(* IEC 61131-3 sources: codesys-framework/txt/application/ToDo/Warnings and Alarms, 15 files *)

(* ---- E_EventLevels.dut.st ---- *)
{attribute 'qualified_only'}
{attribute 'strict'}
TYPE E_EventLevels :
(
	Invalid := 0,
	NotApplicable := 1,
	Success := 5,
	EventIsInformational := 10,
	EventIsWarning_NotUrgent := 20,
	EventIsWarning_Urgent := 21,
	EventIsAlarm_OnlyLogLevel := 40,
	EventIsAlarm_OperatorLevel := 41,
	EventIsAlarm_SupervisorLevel := 42
);
END_TYPE

(* ---- SC_EventConfig.dut.st ---- *)
TYPE SC_EventConfig :
STRUCT
	udiEventID 						: UDINT;
	eSubMachine 					: INT;
	xEventIsDisabled 				: BOOL := FALSE;
	eEventLevel_InCaseOfWarning 	: E_EventLevels;
	eEventLevel_InCaseOfAlarm 		: E_EventLevels;
END_STRUCT
END_TYPE

(* ---- SC_EventHandler.dut.st ---- *)
TYPE SC_EventHandler :
STRUCT
	scEventConfig 					: SC_EventConfig;
	eEventLevel 					: E_EventLevels;
	xEvent_WarningIsActive 			: BOOL;
	xEvent_AlarmIsActive 			: BOOL;
	xEvent_WarningInsertedInLog 	: BOOL;
	xEvent_AlarmInsertedInLog 		: BOOL;
END_STRUCT
END_TYPE

(* ---- F_Event_InsertInLog.pou.st ---- *)
FUNCTION F_Event_InsertInLog : BOOL
VAR_INPUT
	eSubMachine 			: INT;
	w 						: WORD;
	udiEventID 				: UDINT;
	eEventLevel 			: E_EventLevels;
	asEventPayload 			: ARRAY [1..cHYP_MAX_PAYLOADFIELDS] OF STRING;
END_VAR
VAR
	_scEventForHyperion 	: SC_Hyperion_EventStruct;
END_VAR

// --- BEGIN IMPLEMENTATION ---

IF eSubMachine = E_SubMachines.YarnStorage THEN
	audiYSEventCounter[w] := audiYSEventCounter[w] + 1;
	_scEventForHyperion.Counter := audiYSEventCounter[w];

	IF audiYSEventCounter[w] >= 4294967295 THEN
		audiYSEventCounter[w] := 0;
	END_IF

ELSIF eSubMachine = E_SubMachines.CardBoardStorage THEN
	udiCSEventCounter := udiCSEventCounter + 1;
	_scEventForHyperion.Counter := udiCSEventCounter;

	IF udiCSEventCounter >= 4294967295 THEN
		udiCSEventCounter := 0;
	END_IF

ELSE
	udiFREventCounter := udiFREventCounter + 1;
	_scEventForHyperion.Counter := udiFREventCounter;

	IF udiFREventCounter >= 4294967295 THEN
		udiFREventCounter := 0;
	END_IF

END_IF

_scEventForHyperion.Identification := udiEventID;

(*
IF eSubMachine = E_SubMachines.Creel THEN
	audiCLEventCounter[w] := audiCLEventCounter[w] + 1;
	_scEventForHyperion.Counter := audiCLEventCounter[w];
ELSIF eSubMachine = E_SubMachines.CreelRobot THEN
	audiCREventCounter[w] := audiCREventCounter[w] + 1;
	_scEventForHyperion.Counter := audiCREventCounter[w];
ELSIF eSubMachine = E_SubMachines.CreelConveyor THEN
	audiCCEventCounter[w] := audiCCEventCounter[w] + 1;
	_scEventForHyperion.Counter := audiCCEventCounter[w];
ELSIF eSubMachine = E_SubMachines.YarnConsumer THEN
	audiHSEventCounter[w] := audiHSEventCounter[w] + 1;
	_scEventForHyperion.Counter := audiHSEventCounter[w];
ELSE
	udiCUEventCounter := udiCUEventCounter + 1;
	_scEventForHyperion.Counter := udiCUEventCounter;
END_IF
*)

_scEventForHyperion.Identification := udiEventID;

// Create Hyperion Event Struct
CASE (eEventLevel) OF
	E_EventLevels.EventIsInformational : _scEventForHyperion.Level := cHYP_LEVEL_INFORMATIONAL;
	E_EventLevels.Success : _scEventForHyperion.Level := cHYP_LEVEL_BOOKMARK;
	E_EventLevels.EventIsWarning_NotUrgent : _scEventForHyperion.Level := cHYP_LEVEL_WARNING;
	E_EventLevels.EventIsWarning_Urgent : _scEventForHyperion.Level := cHYP_LEVEL_WARNING;
	E_EventLevels.EventIsAlarm_OnlyLogLevel : _scEventForHyperion.Level := cHYP_LEVEL_ERROR;
	E_EventLevels.EventIsAlarm_OperatorLevel : _scEventForHyperion.Level := cHYP_LEVEL_ERROR;
	E_EventLevels.EventIsAlarm_SupervisorLevel : _scEventForHyperion.Level := cHYP_LEVEL_ERROR;
END_CASE

// _scEventForHyperion.TimeStamp := sTimeStamp_Local_AsString;
_scEventForHyperion.TimeStamp := sTimeStamp_UTC_AsString;
_scEventForHyperion.PayLoad := F_HyperionCreatePayloadString (asEventPayload := asEventPayload);

// Insert in local eventbuffer
IF eSubMachine = E_SubMachines.YarnStorage THEN
	audiYSLocalEventPointer[w] := audiYSLocalEventPointer[w] + 1;
	IF audiYSLocalEventPointer[w] > cMaxLocalEvents THEN
		audiYSLocalEventPointer[w] := 1;
	END_IF
	aascYSLocalEventList[w][audiYSLocalEventPointer[w]].udiEventID := udiEventID;
	aascYSLocalEventList[w][audiYSLocalEventPointer[w]].eEventLevel := eEventLevel;

ELSE
	udiFRLocalEventPointer := udiFRLocalEventPointer + 1;
	IF udiFRLocalEventPointer > cMaxLocalEvents THEN
		udiFRLocalEventPointer := 1;
	END_IF
	ascFRLocalEventList[udiFRLocalEventPointer].udiEventID := udiEventID;
	ascFRLocalEventList[udiFRLocalEventPointer].eEventLevel := eEventLevel;
END_IF

// Insert in Hyperion eventbuffer
IF eSubMachine = E_SubMachines.YarnStorage THEN
	aiYSHyperionEventPointer[w] := aiYSHyperionEventPointer[w] + 1;
	IF (aiYSHyperionEventPointer[w] > 50) THEN
		aiYSHyperionEventPointer[w] := 1;
	END_IF
	aascYSHyperion_EventList[w][aiYSHyperionEventPointer[w]] := _scEventForHyperion;
ELSE
	iFRHyperionEventPointer := iFRHyperionEventPointer + 1;
	IF (iFRHyperionEventPointer > cHYP_MAX_EVENTS) THEN
		iFRHyperionEventPointer := 1;
	END_IF
	ascFRHyperion_EventList[iFRHyperionEventPointer] := _scEventForHyperion;
END_IF

(* ---- F_Event_InsertMessage.pou.st ---- *)
FUNCTION F_Event_InsertMessage : BOOL
VAR_INPUT
	eSubMachine : INT;
	w : WORD;
	iComponentID : INT;
	udiEventID : UDINT;
	eEventLevel : E_EventLevels;
END_VAR
VAR
END_VAR
VAR_IN_OUT
END_VAR
VAR
	_asEventPayload : ARRAY [1..10] OF STRING;
	_i : INT;
END_VAR

// --- BEGIN IMPLEMENTATION ---

// Payload
_asEventPayload[1] := INT_TO_STRING (iComponentID);
FOR _i := 2 TO 10 BY 1 DO
	_asEventPayload[_i] := '';
END_FOR

// Insert in log
F_Event_InsertInLog (
	eSubMachine := eSubMachine,
	w := w,
	udiEventID := udiEventID,
	eEventLevel := eEventLevel,
	asEventPayload := _asEventPayload
);

(* ---- F_Event_InsertMessage_ParameterChange.pou.st ---- *)
FUNCTION F_Event_InsertMessage_ParameterChange : BOOL
VAR_INPUT
	eSubMachine : INT;
	w : WORD;
	udiEventID : UDINT;
	eValidationCode : E_ParameterValidationCode;
	rParameterValue_Previous : REAL;
	rParameterValue_New : REAL;
	rParameterValue_MinimumValue : REAL;
	rParameterValue_MaximumValue : REAL;
END_VAR
VAR
	_eEventLevel : E_EventLevels;
	_asEventPayload : ARRAY [1..10] OF STRING;
	_i : INT;
END_VAR

// --- BEGIN IMPLEMENTATION ---

// Parameter
CASE (eValidationCode) OF
	E_ParameterValidationCode.Invalid :
		_asEventPayload[1] := '-';
		_eEventLevel := E_EventLevels.EventIsWarning_Urgent;
	E_ParameterValidationCode.Validation_Failed_IsZero :
		_asEventPayload[1] := '=0';
		_eEventLevel := E_EventLevels.EventIsWarning_Urgent;
	E_ParameterValidationCode.Validation_Failed_BelowMinimum :
		_asEventPayload[1] := '<';
		_eEventLevel := E_EventLevels.EventIsWarning_Urgent;
	E_ParameterValidationCode.Validation_Failed_AboveMaximum :
		_asEventPayload[1] := '>';
		_eEventLevel := E_EventLevels.EventIsWarning_Urgent;
	E_ParameterValidationCode.Validation_Failed_External :
		_asEventPayload[1] := 'Ext';
		_eEventLevel := E_EventLevels.EventIsWarning_Urgent;
	E_ParameterValidationCode.Validation_Ok :
		_asEventPayload[1] := 'V';
		_eEventLevel := E_EventLevels.EventIsInformational;
END_CASE

_asEventPayload[2] := REAL_TO_STRING (rParameterValue_Previous);
_asEventPayload[3] := REAL_TO_STRING (rParameterValue_New);
_asEventPayload[4] := REAL_TO_STRING (rParameterValue_MinimumValue);
_asEventPayload[5] := REAL_TO_STRING (rParameterValue_MaximumValue);

FOR _i := 6 TO 10 BY 1 DO
	_asEventPayload[_i] := '';
END_FOR

F_Event_InsertInLog (
	eSubMachine := eSubMachine,
	w := w,
	udiEventID := udiEventID,
	eEventLevel := _eEventLevel,
	asEventPayload := _asEventPayload
);

(* ---- F_Event_InsertMessage_StringParameterChange.pou.st ---- *)
FUNCTION F_Event_InsertMessage_StringParameterChange : BOOL
VAR_INPUT
	eSubMachine : INT;
	w : WORD;
	udiEventID : UDINT;
	eValidationCode : E_ParameterValidationCode;
	sParameterValue_Previous : STRING;
	sParameterValue_New : STRING;
	iParameterValue_MinimumValue : INT;
	iParameterValue_MaximumValue : INT;
END_VAR
VAR
	_eEventLevel : E_EventLevels;
	_asEventPayload : ARRAY [1..10] OF STRING;
	_i : INT;
END_VAR

// --- BEGIN IMPLEMENTATION ---

//Parameter
CASE (eValidationCode) OF
	E_ParameterValidationCode.Invalid :
		_asEventPayload[1] := '-';
		_eEventLevel := E_EventLevels.EventIsWarning_Urgent;
	E_ParameterValidationCode.Validation_Failed_IsZero :
		_asEventPayload[1] := '=0';
		_eEventLevel := E_EventLevels.EventIsWarning_Urgent;
	E_ParameterValidationCode.Validation_Failed_BelowMinimum :
		_asEventPayload[1] := '<';
		_eEventLevel := E_EventLevels.EventIsWarning_Urgent;
	E_ParameterValidationCode.Validation_Failed_AboveMaximum :
		_asEventPayload[1] := '>';
		_eEventLevel := E_EventLevels.EventIsWarning_Urgent;
	E_ParameterValidationCode.Validation_Failed_External :
		_asEventPayload[1] := 'Ext';
		_eEventLevel := E_EventLevels.EventIsWarning_Urgent;
	E_ParameterValidationCode.Validation_Ok :
		_asEventPayload[1] := 'V';
		_eEventLevel := E_EventLevels.EventIsInformational;
END_CASE

_asEventPayload[2] := sParameterValue_Previous;
_asEventPayload[3] := sParameterValue_New;
_asEventPayload[4] := INT_TO_STRING (iParameterValue_MinimumValue);
_asEventPayload[5] := INT_TO_STRING (iParameterValue_MaximumValue);

FOR _i := 6 TO 10 BY 1 DO
	_asEventPayload[_i] := '';
END_FOR

F_Event_InsertInLog (
	eSubMachine := eSubMachine,
	w := w,
	udiEventID := udiEventID,
	eEventLevel := _eEventLevel,
	asEventPayload := _asEventPayload
);

(* ---- F_Event_InsertMessageComponentID.pou.st ---- *)
FUNCTION F_Event_InsertMessageComponentID : BOOL
VAR_INPUT
	eSubMachine : INT;
	w : WORD;
	iComponentID : INT;
	udiEventID : UDINT;
	eEventLevel : E_EventLevels;
	sMessageString : STRING;
END_VAR
VAR
END_VAR
VAR_IN_OUT
END_VAR
VAR
	_asEventPayload : ARRAY [1..10] OF STRING;
	_i : INT;
END_VAR

// --- BEGIN IMPLEMENTATION ---

// Payload
_asEventPayload[1] := INT_TO_STRING (iComponentID);
_asEventPayload[2] := sMessageString;
FOR _i := 3 TO 10 BY 1 DO
	_asEventPayload[_i] := '';
END_FOR

// Insert in log
F_Event_InsertInLog (
	eSubMachine := eSubMachine,
	w := w,
	udiEventID := udiEventID,
	eEventLevel := eEventLevel,
	asEventPayload := _asEventPayload
);

(* ---- F_Event_InsertMessageString.pou.st ---- *)
FUNCTION F_Event_InsertMessageString : BOOL
VAR_INPUT
	eSubMachine 		: INT;
	w 					: WORD;
	udiEventID 			: UDINT;
	eEventLevel 		: E_EventLevels;
	sMessageString1 	: STRING;
	sMessageString2 	: STRING;
END_VAR
VAR
END_VAR
VAR_IN_OUT
END_VAR
VAR
	_asEventPayload 	: ARRAY[1..10] OF STRING;
	_i 					: INT;
END_VAR

// --- BEGIN IMPLEMENTATION ---

// Payload
_asEventPayload[1] := sMessageString1;
_asEventPayload[2] := sMessageString2;

FOR _i := 3 TO 10 BY 1 DO
	_asEventPayload[_i] := '';
END_FOR

// Insert in log
F_Event_InsertInLog (
	eSubMachine := eSubMachine,
	w := w,
	udiEventID := udiEventID,
	eEventLevel := eEventLevel,
	asEventPayload := _asEventPayload
);

(* ---- F_Event_InsertPLCEventRqst.pou.st ---- *)
FUNCTION F_Event_InsertPLCEventRqst : BOOL
VAR_INPUT
	eSubMachine : INT;
	w : WORD;
	udiEventID : UDINT;
END_VAR
VAR
END_VAR
VAR_IN_OUT
END_VAR
VAR
	_asEventPayload : ARRAY[1..10] OF STRING;
	_i : int;
END_VAR

// --- BEGIN IMPLEMENTATION ---

//Payload
_asEventPayload[1] := ' TEST';
FOR _i := 2 TO 10 BY 1 DO
	_asEventPayload[_i] := '';
END_FOR

//Insert in log
F_Event_InsertInLog(
	eSubMachine := eSubMachine,
	w := w,
	udiEventID := udiEventID,
	eEventLevel := E_EventLevels.EventIsInformational,
	asEventPayload := _asEventPayload
);

(* ---- F_Event_InsertPLCServiceRqst.pou.st ---- *)
FUNCTION F_Event_InsertPLCServiceRqst : BOOL
VAR_INPUT
	eSubMachine : INT;
	w : WORD;
	udiEventID : UDINT;
	iPLCServiceRqst : INT;
END_VAR
VAR
END_VAR
VAR_IN_OUT
END_VAR
VAR
	_asEventPayload : ARRAY [1..10] OF STRING;
	_i : INT;
END_VAR

// --- BEGIN IMPLEMENTATION ---

// Payload
_asEventPayload[1] := INT_TO_STRING (iPLCServiceRqst);
FOR _i := 2 TO 10 BY 1 DO
	_asEventPayload[_i] := '';
END_FOR

// Insert in log
F_Event_InsertInLog (
	eSubMachine := eSubMachine,
	w := w,
	udiEventID := udiEventID,
	eEventLevel := E_EventLevels.EventIsInformational,
	asEventPayload := _asEventPayload
);

(* ---- F_EventHandler_AnalogLevelMonitor.pou.st ---- *)
FUNCTION F_EventHandler_AnalogLevelMonitor : BOOL
VAR_INPUT
	eSubMachine : INT;
	w : WORD;
	iComponentId : INT;
	rProcessValue : REAL;
	rAlarmLevelLow : REAL;
	rWarningLevelLow : REAL;
	rWarningLevelHigh : REAL;
	rAlarmLevelHigh : REAL;
	xReset : BOOL;
	xAlarmHigh : BOOL;
	xWarningHigh : BOOL;
	xWarningLow : BOOL;
	xAlarmLow : BOOL;
END_VAR
VAR
END_VAR
VAR_IN_OUT
	scEvent : SC_EventHandler;
END_VAR
VAR
	_asEventPayload : ARRAY [1..10] OF STRING;
	_i : INT;
END_VAR

// --- BEGIN IMPLEMENTATION ---

// Reset
IF xReset THEN
	scEvent.xEvent_WarningInsertedInLog := FALSE;
	scEvent.xEvent_AlarmInsertedInLog := FALSE;
	RETURN;
END_IF

// Check disabled
IF scEvent.scEventConfig.xEventIsDisabled THEN
	scEvent.xEvent_WarningInsertedInLog := FALSE;
	scEvent.xEvent_AlarmInsertedInLog := FALSE;
	RETURN;
END_IF

// Insert in log - Warning
IF scEvent.xEvent_WarningIsActive AND NOT scEvent.xEvent_WarningInsertedInLog THEN
	// Payload
	_asEventPayload[1] := INT_TO_STRING (iComponentID);
	_asEventPayload[2] := REAL_TO_STRING (rProcessValue);
	_asEventPayload[3] := REAL_TO_STRING (rAlarmLevelLow);
	_asEventPayload[4] := REAL_TO_STRING (rWarningLevelLow);
	_asEventPayload[5] := REAL_TO_STRING (rWarningLevelHigh);
	_asEventPayload[6] := REAL_TO_STRING (rAlarmLevelHigh);

	IF xAlarmHigh THEN
	_asEventPayload[7] := 'Alarm HIGH tension';
	ELSIF xAlarmLow THEN
	_asEventPayload[7] := 'Alarm LOW tension';
	ELSIF xWarningHigh THEN
	_asEventPayload[7] := 'Warning HIGH tension';
	ELSIF xWarningLow THEN
	_asEventPayload[7] := 'Warning LOW tension';
	END_IF

	FOR _i := 8 TO 10 BY 1 DO
		_asEventPayload[_i] := '';
	END_FOR
	F_Event_InsertInLog (
		eSubMachine := eSubMachine,
		w := w,
		udiEventID := scEvent.scEventConfig.udiEventID,
		eEventLevel := scEvent.scEventConfig.eEventLevel_InCaseOfWarning,
		asEventPayload := _asEventPayload
	);
	scEvent.xEvent_WarningInsertedInLog := TRUE;
END_IF

// Insert in log - Alarm
IF scEvent.xEvent_AlarmIsActive AND NOT scEvent.xEvent_AlarmInsertedInLog THEN
	// Payload
	_asEventPayload[1] := INT_TO_STRING (iComponentID);
	_asEventPayload[2] := REAL_TO_STRING (rProcessValue);
	_asEventPayload[3] := REAL_TO_STRING (rAlarmLevelLow);
	_asEventPayload[4] := REAL_TO_STRING (rWarningLevelLow);
	_asEventPayload[5] := REAL_TO_STRING (rWarningLevelHigh);
	_asEventPayload[6] := REAL_TO_STRING (rAlarmLevelHigh);

	IF xAlarmHigh THEN
	_asEventPayload[7] := 'Alarm HIGH tension';
	ELSIF xAlarmLow THEN
	_asEventPayload[7] := 'Alarm LOW tension';
	ELSIF xWarningHigh THEN
	_asEventPayload[7] := 'Warning HIGH tension';
	ELSIF xWarningLow THEN
	_asEventPayload[7] := 'Warning LOW tension';
	ELSE
	_asEventPayload[7] := '';
	END_IF

	FOR _i := 8 TO 10 BY 1 DO
		_asEventPayload[_i] := '';
	END_FOR
	F_Event_InsertInLog (
		eSubMachine := eSubMachine,
		w := w,
		udiEventID := scEvent.scEventConfig.udiEventID,
		eEventLevel := scEvent.scEventConfig.eEventLevel_InCaseOfAlarm,
		asEventPayload := _asEventPayload
	);
	scEvent.xEvent_AlarmInsertedInLog := TRUE;
END_IF

(* ---- F_EventHandler_Component.pou.st ---- *)
FUNCTION F_EventHandler_Component : BOOL
VAR_INPUT
	eSubMachine : INT;
	w : WORD;
	iComponentId : INT;
	sComponentName : STRING;//STRING [10];
	xReset : BOOL;
END_VAR
VAR
END_VAR
VAR_IN_OUT
	scEvent : SC_EventHandler;
END_VAR
VAR
	_asEventPayload : ARRAY [1..10] OF STRING;
	_i : INT;
END_VAR

// --- BEGIN IMPLEMENTATION ---

// Check disabled
IF scEvent.scEventConfig.xEventIsDisabled THEN
	scEvent.xEvent_WarningInsertedInLog := FALSE;
	scEvent.xEvent_AlarmInsertedInLog := FALSE;
	RETURN;
END_IF

// Insert in log
IF scEvent.xEvent_WarningIsActive AND NOT scEvent.xEvent_WarningInsertedInLog OR
	scEvent.xEvent_AlarmIsActive AND NOT scEvent.xEvent_AlarmInsertedInLog
THEN
	// Payload
	_asEventPayload[1] := INT_TO_STRING (iComponentId);
	_asEventPayload[2] := sComponentName;

	FOR _i := 3 TO 10 BY 1 DO
		_asEventPayload[_i] := '';
	END_FOR

	IF scEvent.xEvent_AlarmIsActive THEN

		F_Event_InsertInLog (
			eSubMachine := eSubMachine,
			w := w,
			udiEventID := scEvent.scEventConfig.udiEventID,
			eEventLevel := scEvent.scEventConfig.eEventLevel_InCaseOfAlarm,
			asEventPayload := _asEventPayload
		);

	ELSE

		F_Event_InsertInLog (
			eSubMachine := eSubMachine,
			w := w,
			udiEventID := scEvent.scEventConfig.udiEventID,
			eEventLevel := scEvent.scEventConfig.eEventLevel_InCaseOfWarning,
			asEventPayload := _asEventPayload
		);

	END_IF

	IF scEvent.xEvent_AlarmIsActive THEN
		scEvent.xEvent_AlarmInsertedInLog := TRUE;
	ELSE
		scEvent.xEvent_WarningInsertedInLog := TRUE;
	END_IF
END_IF

(* ---- F_EventHandler_Component_RaiseEvent.pou.st ---- *)
FUNCTION F_EventHandler_Component_RaiseEvent : BOOL
VAR_INPUT
	w : WORD;
	iComponentId : INT;
	sComponentName : STRING;//STRING [10];
END_VAR
VAR
END_VAR
VAR_IN_OUT
	scEvent : SC_EventHandler;
END_VAR
VAR
	_asEventPayload : ARRAY [1..10] OF STRING;
	_i : INT;
END_VAR

// --- BEGIN IMPLEMENTATION ---

// Check disabled
IF scEvent.scEventConfig.xEventIsDisabled THEN
	scEvent.xEvent_WarningInsertedInLog := FALSE;
	scEvent.xEvent_AlarmInsertedInLog := FALSE;
	RETURN;
END_IF

// Insert in log
IF scEvent.xEvent_WarningIsActive AND NOT scEvent.xEvent_WarningInsertedInLog OR
	scEvent.xEvent_AlarmIsActive AND NOT scEvent.xEvent_AlarmInsertedInLog
THEN
	// Payload
	_asEventPayload[1] := INT_TO_STRING (iComponentId);
	_asEventPayload[2] := sComponentName;

	FOR _i := 3 TO 10 BY 1 DO
		_asEventPayload[_i] := '';
	END_FOR

	IF scEvent.xEvent_AlarmIsActive THEN

		F_Event_InsertInLog (
			eSubMachine := scEvent.scEventConfig.eSubMachine,
			w := w,
			udiEventID := scEvent.scEventConfig.udiEventID,
			eEventLevel := scEvent.scEventConfig.eEventLevel_InCaseOfAlarm,
			asEventPayload := _asEventPayload
		);

	ELSE

		F_Event_InsertInLog (
			eSubMachine := scEvent.scEventConfig.eSubMachine,
			w := w,
			udiEventID := scEvent.scEventConfig.udiEventID,
			eEventLevel := scEvent.scEventConfig.eEventLevel_InCaseOfWarning,
			asEventPayload := _asEventPayload
		);

	END_IF

	IF scEvent.xEvent_AlarmIsActive THEN
		scEvent.xEvent_AlarmInsertedInLog := TRUE;
	ELSE
		scEvent.xEvent_WarningInsertedInLog := TRUE;
	END_IF

END_IF

(* ---- F_HyperionCreatePayloadString.pou.st ---- *)
FUNCTION F_HyperionCreatePayloadString : ARRAY[0..63] OF BYTE
VAR_INPUT
	asEventPayload : ARRAY[1..10] OF STRING;
END_VAR
VAR
	_sSeparator : STRING(1);
	_bySeparatorAsciiValue : BYTE;
	_byCharAsciiValue : BYTE;
	_iCounter : INT;
	_sPayloadPartString : STRING;
	_sPayloadString : STRING (cHYP_MAX_PAYLOADBYTESIZE);
	_iPayloadStringLength : INT;

	_abyPayloadByteArray : POINTER TO ARRAY [0 .. cHYP_MAX_PAYLOADBYTESIZE] OF BYTE;
	_abyPayloadByteArray_Return : ARRAY [0 .. cHYP_MAX_PAYLOADBYTESIZE] OF BYTE;
END_VAR

// --- BEGIN IMPLEMENTATION ---

// Init
_sPayloadString := '';
_sSeparator := ';';
_bySeparatorAsciiValue := 59;
// Check PayloadStrings
FOR _iCounter := 1 TO cHYP_MAX_PAYLOADFIELDS BY 1 DO

	IF asEventPayload[_iCounter] = '' THEN
		EXIT;
	END_IF

	_sPayloadPartString := CONCAT(STR1 := asEventPayload[_iCounter], STR2 := _sSeparator);
	_sPayloadString := CONCAT(STR1 := _sPayloadString, STR2 := _sPayloadPartString);
END_FOR

// String to ByteArray
_iPayloadStringLength := LEN (STR := _sPayloadString);
_abyPayloadByteArray := ADR (_sPayloadString);

// Replace ';' with 0
FOR _iCounter := 0 TO cHYP_MAX_PAYLOADBYTESIZE BY 1 DO
	IF _iCounter < _iPayloadStringLength THEN
		_byCharAsciiValue := _abyPayloadByteArray^[_iCounter];
 		IF (_byCharAsciiValue <> _bySeparatorAsciiValue) THEN
			_abyPayloadByteArray_Return[_iCounter] := _byCharAsciiValue;
		ELSE
			_abyPayloadByteArray_Return[_iCounter] := 0;
		END_IF
	ELSE
		_abyPayloadByteArray_Return[_iCounter] := 0;
	END_IF
END_FOR

F_HyperionCreatePayloadString := _abyPayloadByteArray_Return;
